Fanuc KAREL source: KA00030.KL

PROGRAM KA00030
%NOLOCKGROUP
VAR
  SRC: BOOLEAN
  DST: XYZWPR
BEGIN
  SRC = TRUE
  DST = SRC
END KA00030
